FUNCTION_BLOCK FB_MotionSystem
VAR
    fbXPlanarSystem   : FB_XPlanarSystem;
    fbXPlanarMover    : ARRAY[1..maxNumMover] OF FB_XPlanarMoverStandard;
    nStartupSequence  : UDINT;
    nStartingSequence : UDINT;
END_VAR

METHOD Cycle
VAR
    i : UDINT;
END_VAR
// Call every PLC cycle: updates the XPlanar system and the movers.
fbXPlanarSystem.Cycle();
FOR i := 1 TO moverCount DO
    fbXPlanarMover[i].Cycle();
END_FOR
END_METHOD

METHOD Startup : BOOL
VAR
    i : UDINT;
END_VAR
// One-time setup: register movers (and tracks) in the system. TRUE when done.
CASE nStartupSequence OF
    0:  nStartupSequence := 1;
    1:  FOR i := 1 TO moverCount DO
            fbXPlanarSystem.SetMoverStandard(i, fbXPlanarMover[i]);
        END_FOR
        nStartupSequence := 30;
    30: Startup := TRUE;
END_CASE
END_METHOD

METHOD Starting : BOOL
VAR_INPUT
    bReset : BOOL;
END_VAR
// Brings the system to a ready state step by step. TRUE when done.
IF bReset THEN
    Starting := FALSE;
    nStartingSequence := 0;
END_IF
CASE nStartingSequence OF
    // start
    0:  nStartingSequence := 50;
    // enable movers
    50: IF fbXPlanarSystem.EnableMovers() THEN
            nStartingSequence := 51;
        END_IF
    // wait for enable
    51: IF fbXPlanarSystem.P_EnableMovers.Done THEN
            nStartingSequence := 80;
        ELSIF fbXPlanarSystem.P_EnableMovers.Error THEN
            nStartingSequence := 90;   // enable failed
        END_IF
    // ready
    80: Starting := TRUE;
END_CASE
END_METHOD

END_FUNCTION_BLOCK

(* stored: Version 1.1.0.1
   POU FB_MotionSystem: Id {76b90533-2f5f-4265-a888-7463c8f15552}, SpecialFunc None
   Method Cycle: Id {7a6a436f-abe3-49cf-80ba-736989644d1a}
   Method Startup: Id {ab1988d1-2b56-4e22-9706-835668cd8a23}
   Method Starting: Id {04721e65-d0d5-4973-a78a-e55f3a27c0da} *)
